Universal Robots PolyScope program: TgtProg.urp

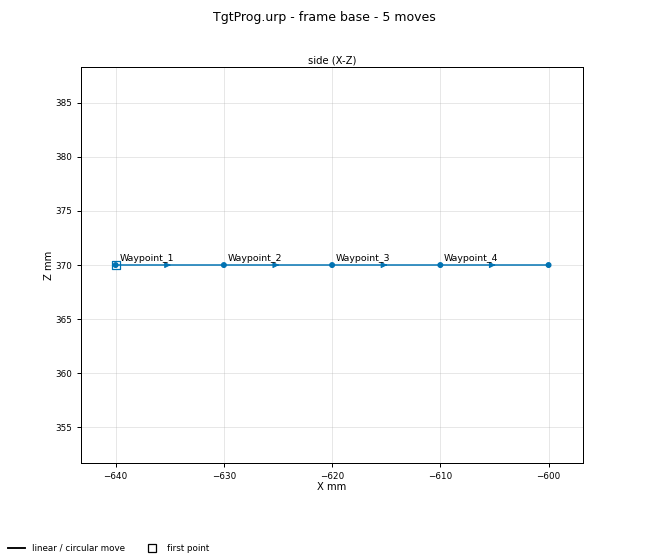
[picture p0: tool path of TgtProg.urp in frame base, 5 of 5 moves have a stored position in this frame; points joined in program order, loops and branches not executed]
Program TgtProg (createdIn=3.0.0 lastSavedIn=3.0.0 directory=/programs installation=default)
Robot Program (runOnlyOnce=true motionType=MoveJ speed=1.047198 acceleration=1.396263 useActiveTCP=false)
  'Program generated by RoboDK v6.0.7 for UR10 on XX/XX/XXXX 18:00:00'
  'Using nominal kinematics.'
  MoveL speed 250 mm/s, acceleration 1200 mm/s^2 (useActiveTCP=true)
    Waypoint Waypoint_1: TCP in base x=-640 y=500 z=370 mm, rx=0.732 ry=2.1859 rz=-0.5703 rad; joints [0, -10, 20, 0, 30, 0] deg
    Waypoint Waypoint_2: TCP in base x=-630 y=500 z=370 mm, rx=0.732 ry=2.1859 rz=-0.5703 rad; joints [0, -10, 20, 0, 30, 0] deg
    Waypoint Waypoint_3: TCP in base x=-620 y=500 z=370 mm, rx=0.732 ry=2.1859 rz=-0.5703 rad; joints [0, -10, 20, 0, 30, 0] deg
    Waypoint Waypoint_4: TCP in base x=-610 y=500 z=370 mm, rx=0.732 ry=2.1859 rz=-0.5703 rad; joints [0, -10, 20, 0, 30, 0] deg
    Waypoint Waypoint_5: TCP in base x=-600 y=500 z=370 mm, rx=0.732 ry=2.1859 rz=-0.5703 rad; joints [0, -10, 20, 0, 30, 0] deg
